// TIA Portal V20 export
// export: Created 2026-10-12T16:46:19.999098Z, ExportSetting WithDefaults, DisplayName Totally Integrated Automation Portal, DisplayVersion V20 Update 6, DisplayName TIA Portal Openness, DisplayVersion V20 Update 6, DisplayName TIA Portal Version Control Interface, DisplayVersion V20 Update 6, DisplayName SINAMICS Startdrive Advanced, DisplayVersion V20 SP1 Update 2, DisplayName SINAMICS Startdrive G110M, G120, G120C, G120D, G120P, G115D, DisplayVersion V20 SP1 Update 2, DisplayName SINAMICS Startdrive G130, G150, S120, S150, SINAMICS MV, G220, S200, S210, DisplayVersion V20 SP1 Update 2, DisplayName STEP 7 Professional, DisplayVersion V20 Update 6, DisplayName STEP 7 Safety, DisplayVersion V20 Update 2, DisplayName WinCC Basic/Comfort/Advanced, DisplayVersion V20 Update 6, DisplayName WinCC Professional, DisplayVersion V20 Update 6, DisplayName WinCC Unified, DisplayVersion V20 Update 6
DATA_BLOCK "DB_FlexKraft_Data"   // DB5
{ S7_Optimized_Access := 'FALSE' }
VERSION : 0.1
// ==============================================================================
//  DB: Daten aller drei FlexKraft-GerÃ¤te
// ==============================================================================
// stored: AutoNumber true, DBAccessibleFromOPCUA true, DBAccessibleFromWebserver true, IsOnlyStoredInLoadMemory false, IsWriteProtectedInAS false
   VAR
      FK_1 { S7_SetPoint := 'True'} : "UDT_FlexKraft_Device";   // ModbusAdr 2 (Gateway-Bytes 0..31)
      FK_2 { S7_SetPoint := 'True'} : "UDT_FlexKraft_Device";   // ModbusAdr 3 (Gateway-Bytes 32..63)
      FK_3 { S7_SetPoint := 'True'} : "UDT_FlexKraft_Device";   // ModbusAdr 4 (Gateway-Bytes 64..95)
   END_VAR
BEGIN
END_DATA_BLOCK
